(* IEC 61131-3 sources: STAR-PLC-Agent/results/raw/four_group_20261114/star_terra/PUB009/generation/sim_00, 1 file *)

(* ---- test_program.st ---- *)
PROGRAM PLC_PRG
VAR
 BenchStep : UDINT := 0;
 BenchCalls : UDINT := 0;
 BenchDone : BOOL := FALSE;
 BenchUut0 : FB_Task;
 BenchUut1 : FB_Task;
 TraceIn_cyclicExecution : ARRAY[0..15] OF BOOL;
 TraceIn_trigger : ARRAY[0..15] OF BOOL;
 TraceIn_value : ARRAY[0..15] OF LREAL;
 TraceIn_windowSize : ARRAY[0..15] OF INT;
 TraceIn_reset : ARRAY[0..15] OF BOOL;
 TraceOut_average : ARRAY[0..15] OF LREAL;
 TraceOut_windowSizeReached : ARRAY[0..15] OF BOOL;
 TraceOut_error : ARRAY[0..15] OF BOOL;
 TraceOut_status : ARRAY[0..15] OF WORD;
END_VAR

IF NOT BenchDone THEN
 CASE BenchStep OF
 0:
   BenchUut0.cyclicExecution := FALSE;
   BenchUut0.trigger := FALSE;
   BenchUut0.value := LREAL#100.0;
   BenchUut0.windowSize := INT#3;
   BenchUut0.reset := FALSE;
   TraceIn_cyclicExecution[0] := BenchUut0.cyclicExecution;
   TraceIn_trigger[0] := BenchUut0.trigger;
   TraceIn_value[0] := BenchUut0.value;
   TraceIn_windowSize[0] := BenchUut0.windowSize;
   TraceIn_reset[0] := BenchUut0.reset;
   BenchUut0();
   TraceOut_average[0] := BenchUut0.average;
   TraceOut_windowSizeReached[0] := BenchUut0.windowSizeReached;
   TraceOut_error[0] := BenchUut0.error;
   TraceOut_status[0] := BenchUut0.status;
   BenchCalls := BenchCalls + 1;
 1:
   BenchUut0.cyclicExecution := FALSE;
   BenchUut0.trigger := TRUE;
   BenchUut0.value := LREAL#3.0;
   BenchUut0.windowSize := INT#3;
   BenchUut0.reset := FALSE;
   TraceIn_cyclicExecution[1] := BenchUut0.cyclicExecution;
   TraceIn_trigger[1] := BenchUut0.trigger;
   TraceIn_value[1] := BenchUut0.value;
   TraceIn_windowSize[1] := BenchUut0.windowSize;
   TraceIn_reset[1] := BenchUut0.reset;
   BenchUut0();
   TraceOut_average[1] := BenchUut0.average;
   TraceOut_windowSizeReached[1] := BenchUut0.windowSizeReached;
   TraceOut_error[1] := BenchUut0.error;
   TraceOut_status[1] := BenchUut0.status;
   BenchCalls := BenchCalls + 1;
 2:
   BenchUut0.cyclicExecution := FALSE;
   BenchUut0.trigger := TRUE;
   BenchUut0.value := LREAL#99.0;
   BenchUut0.windowSize := INT#3;
   BenchUut0.reset := FALSE;
   TraceIn_cyclicExecution[2] := BenchUut0.cyclicExecution;
   TraceIn_trigger[2] := BenchUut0.trigger;
   TraceIn_value[2] := BenchUut0.value;
   TraceIn_windowSize[2] := BenchUut0.windowSize;
   TraceIn_reset[2] := BenchUut0.reset;
   BenchUut0();
   TraceOut_average[2] := BenchUut0.average;
   TraceOut_windowSizeReached[2] := BenchUut0.windowSizeReached;
   TraceOut_error[2] := BenchUut0.error;
   TraceOut_status[2] := BenchUut0.status;
   BenchCalls := BenchCalls + 1;
 3:
   BenchUut0.cyclicExecution := TRUE;
   BenchUut0.trigger := FALSE;
   BenchUut0.value := LREAL#6.0;
   BenchUut0.windowSize := INT#3;
   BenchUut0.reset := FALSE;
   TraceIn_cyclicExecution[3] := BenchUut0.cyclicExecution;
   TraceIn_trigger[3] := BenchUut0.trigger;
   TraceIn_value[3] := BenchUut0.value;
   TraceIn_windowSize[3] := BenchUut0.windowSize;
   TraceIn_reset[3] := BenchUut0.reset;
   BenchUut0();
   TraceOut_average[3] := BenchUut0.average;
   TraceOut_windowSizeReached[3] := BenchUut0.windowSizeReached;
   TraceOut_error[3] := BenchUut0.error;
   TraceOut_status[3] := BenchUut0.status;
   BenchCalls := BenchCalls + 1;
 4:
   BenchUut0.cyclicExecution := TRUE;
   BenchUut0.trigger := TRUE;
   BenchUut0.value := LREAL#9.0;
   BenchUut0.windowSize := INT#3;
   BenchUut0.reset := FALSE;
   TraceIn_cyclicExecution[4] := BenchUut0.cyclicExecution;
   TraceIn_trigger[4] := BenchUut0.trigger;
   TraceIn_value[4] := BenchUut0.value;
   TraceIn_windowSize[4] := BenchUut0.windowSize;
   TraceIn_reset[4] := BenchUut0.reset;
   BenchUut0();
   TraceOut_average[4] := BenchUut0.average;
   TraceOut_windowSizeReached[4] := BenchUut0.windowSizeReached;
   TraceOut_error[4] := BenchUut0.error;
   TraceOut_status[4] := BenchUut0.status;
   BenchCalls := BenchCalls + 1;
 5:
   BenchUut0.cyclicExecution := FALSE;
   BenchUut0.trigger := TRUE;
   BenchUut0.value := LREAL#99.0;
   BenchUut0.windowSize := INT#3;
   BenchUut0.reset := FALSE;
   TraceIn_cyclicExecution[5] := BenchUut0.cyclicExecution;
   TraceIn_trigger[5] := BenchUut0.trigger;
   TraceIn_value[5] := BenchUut0.value;
   TraceIn_windowSize[5] := BenchUut0.windowSize;
   TraceIn_reset[5] := BenchUut0.reset;
   BenchUut0();
   TraceOut_average[5] := BenchUut0.average;
   TraceOut_windowSizeReached[5] := BenchUut0.windowSizeReached;
   TraceOut_error[5] := BenchUut0.error;
   TraceOut_status[5] := BenchUut0.status;
   BenchCalls := BenchCalls + 1;
 6:
   BenchUut0.cyclicExecution := FALSE;
   BenchUut0.trigger := FALSE;
   BenchUut0.value := LREAL#99.0;
   BenchUut0.windowSize := INT#3;
   BenchUut0.reset := FALSE;
   TraceIn_cyclicExecution[6] := BenchUut0.cyclicExecution;
   TraceIn_trigger[6] := BenchUut0.trigger;
   TraceIn_value[6] := BenchUut0.value;
   TraceIn_windowSize[6] := BenchUut0.windowSize;
   TraceIn_reset[6] := BenchUut0.reset;
   BenchUut0();
   TraceOut_average[6] := BenchUut0.average;
   TraceOut_windowSizeReached[6] := BenchUut0.windowSizeReached;
   TraceOut_error[6] := BenchUut0.error;
   TraceOut_status[6] := BenchUut0.status;
   BenchCalls := BenchCalls + 1;
 7:
   BenchUut0.cyclicExecution := FALSE;
   BenchUut0.trigger := TRUE;
   BenchUut0.value := LREAL#12.0;
   BenchUut0.windowSize := INT#3;
   BenchUut0.reset := FALSE;
   TraceIn_cyclicExecution[7] := BenchUut0.cyclicExecution;
   TraceIn_trigger[7] := BenchUut0.trigger;
   TraceIn_value[7] := BenchUut0.value;
   TraceIn_windowSize[7] := BenchUut0.windowSize;
   TraceIn_reset[7] := BenchUut0.reset;
   BenchUut0();
   TraceOut_average[7] := BenchUut0.average;
   TraceOut_windowSizeReached[7] := BenchUut0.windowSizeReached;
   TraceOut_error[7] := BenchUut0.error;
   TraceOut_status[7] := BenchUut0.status;
   BenchCalls := BenchCalls + 1;
 8:
   BenchUut1.cyclicExecution := TRUE;
   BenchUut1.trigger := FALSE;
   BenchUut1.value := LREAL#8.0;
   BenchUut1.windowSize := INT#1;
   BenchUut1.reset := FALSE;
   TraceIn_cyclicExecution[8] := BenchUut1.cyclicExecution;
   TraceIn_trigger[8] := BenchUut1.trigger;
   TraceIn_value[8] := BenchUut1.value;
   TraceIn_windowSize[8] := BenchUut1.windowSize;
   TraceIn_reset[8] := BenchUut1.reset;
   BenchUut1();
   TraceOut_average[8] := BenchUut1.average;
   TraceOut_windowSizeReached[8] := BenchUut1.windowSizeReached;
   TraceOut_error[8] := BenchUut1.error;
   TraceOut_status[8] := BenchUut1.status;
   BenchCalls := BenchCalls + 1;
 9:
   BenchUut1.cyclicExecution := TRUE;
   BenchUut1.trigger := TRUE;
   BenchUut1.value := LREAL#99.0;
   BenchUut1.windowSize := INT#0;
   BenchUut1.reset := TRUE;
   TraceIn_cyclicExecution[9] := BenchUut1.cyclicExecution;
   TraceIn_trigger[9] := BenchUut1.trigger;
   TraceIn_value[9] := BenchUut1.value;
   TraceIn_windowSize[9] := BenchUut1.windowSize;
   TraceIn_reset[9] := BenchUut1.reset;
   BenchUut1();
   TraceOut_average[9] := BenchUut1.average;
   TraceOut_windowSizeReached[9] := BenchUut1.windowSizeReached;
   TraceOut_error[9] := BenchUut1.error;
   TraceOut_status[9] := BenchUut1.status;
   BenchCalls := BenchCalls + 1;
 10:
   BenchUut1.cyclicExecution := FALSE;
   BenchUut1.trigger := TRUE;
   BenchUut1.value := LREAL#50.0;
   BenchUut1.windowSize := INT#1;
   BenchUut1.reset := FALSE;
   TraceIn_cyclicExecution[10] := BenchUut1.cyclicExecution;
   TraceIn_trigger[10] := BenchUut1.trigger;
   TraceIn_value[10] := BenchUut1.value;
   TraceIn_windowSize[10] := BenchUut1.windowSize;
   TraceIn_reset[10] := BenchUut1.reset;
   BenchUut1();
   TraceOut_average[10] := BenchUut1.average;
   TraceOut_windowSizeReached[10] := BenchUut1.windowSizeReached;
   TraceOut_error[10] := BenchUut1.error;
   TraceOut_status[10] := BenchUut1.status;
   BenchCalls := BenchCalls + 1;
 11:
   BenchUut1.cyclicExecution := TRUE;
   BenchUut1.trigger := FALSE;
   BenchUut1.value := LREAL#20.0;
   BenchUut1.windowSize := INT#100;
   BenchUut1.reset := FALSE;
   TraceIn_cyclicExecution[11] := BenchUut1.cyclicExecution;
   TraceIn_trigger[11] := BenchUut1.trigger;
   TraceIn_value[11] := BenchUut1.value;
   TraceIn_windowSize[11] := BenchUut1.windowSize;
   TraceIn_reset[11] := BenchUut1.reset;
   BenchUut1();
   TraceOut_average[11] := BenchUut1.average;
   TraceOut_windowSizeReached[11] := BenchUut1.windowSizeReached;
   TraceOut_error[11] := BenchUut1.error;
   TraceOut_status[11] := BenchUut1.status;
   BenchCalls := BenchCalls + 1;
 12:
   BenchUut1.cyclicExecution := TRUE;
   BenchUut1.trigger := TRUE;
   BenchUut1.value := LREAL#99.0;
   BenchUut1.windowSize := INT#100;
   BenchUut1.reset := TRUE;
   TraceIn_cyclicExecution[12] := BenchUut1.cyclicExecution;
   TraceIn_trigger[12] := BenchUut1.trigger;
   TraceIn_value[12] := BenchUut1.value;
   TraceIn_windowSize[12] := BenchUut1.windowSize;
   TraceIn_reset[12] := BenchUut1.reset;
   BenchUut1();
   TraceOut_average[12] := BenchUut1.average;
   TraceOut_windowSizeReached[12] := BenchUut1.windowSizeReached;
   TraceOut_error[12] := BenchUut1.error;
   TraceOut_status[12] := BenchUut1.status;
   BenchCalls := BenchCalls + 1;
 13:
   BenchUut1.cyclicExecution := FALSE;
   BenchUut1.trigger := TRUE;
   BenchUut1.value := LREAL#50.0;
   BenchUut1.windowSize := INT#100;
   BenchUut1.reset := FALSE;
   TraceIn_cyclicExecution[13] := BenchUut1.cyclicExecution;
   TraceIn_trigger[13] := BenchUut1.trigger;
   TraceIn_value[13] := BenchUut1.value;
   TraceIn_windowSize[13] := BenchUut1.windowSize;
   TraceIn_reset[13] := BenchUut1.reset;
   BenchUut1();
   TraceOut_average[13] := BenchUut1.average;
   TraceOut_windowSizeReached[13] := BenchUut1.windowSizeReached;
   TraceOut_error[13] := BenchUut1.error;
   TraceOut_status[13] := BenchUut1.status;
   BenchCalls := BenchCalls + 1;
 14:
   BenchUut1.cyclicExecution := TRUE;
   BenchUut1.trigger := FALSE;
   BenchUut1.value := LREAL#30.0;
   BenchUut1.windowSize := INT#100;
   BenchUut1.reset := FALSE;
   TraceIn_cyclicExecution[14] := BenchUut1.cyclicExecution;
   TraceIn_trigger[14] := BenchUut1.trigger;
   TraceIn_value[14] := BenchUut1.value;
   TraceIn_windowSize[14] := BenchUut1.windowSize;
   TraceIn_reset[14] := BenchUut1.reset;
   BenchUut1();
   TraceOut_average[14] := BenchUut1.average;
   TraceOut_windowSizeReached[14] := BenchUut1.windowSizeReached;
   TraceOut_error[14] := BenchUut1.error;
   TraceOut_status[14] := BenchUut1.status;
   BenchCalls := BenchCalls + 1;
 15:
   BenchUut1.cyclicExecution := TRUE;
   BenchUut1.trigger := TRUE;
   BenchUut1.value := LREAL#100.0;
   BenchUut1.windowSize := INT#101;
   BenchUut1.reset := TRUE;
   TraceIn_cyclicExecution[15] := BenchUut1.cyclicExecution;
   TraceIn_trigger[15] := BenchUut1.trigger;
   TraceIn_value[15] := BenchUut1.value;
   TraceIn_windowSize[15] := BenchUut1.windowSize;
   TraceIn_reset[15] := BenchUut1.reset;
   BenchUut1();
   TraceOut_average[15] := BenchUut1.average;
   TraceOut_windowSizeReached[15] := BenchUut1.windowSizeReached;
   TraceOut_error[15] := BenchUut1.error;
   TraceOut_status[15] := BenchUut1.status;
   BenchCalls := BenchCalls + 1;
 END_CASE;
 BenchStep := BenchStep + 1;
 IF BenchStep >= 16 THEN BenchDone := TRUE; END_IF;
END_IF;
END_PROGRAM
